FUNCTION_BLOCK FB_AliasLevel2
VAR
    {attribute 'pytmc' := '
        pv:
    '}
    stAlias : ST_Alias;
END_VAR

END_FUNCTION_BLOCK

(* stored: Version 1.1.0.1
   POU FB_AliasLevel2: Id {eea0d705-aed2-40eb-934c-5adef550e14c}, SpecialFunc None *)
